// TIA Portal V20 export
// export: Created 2026-10-20T18:55:29.0460085Z, ExportSetting None, DisplayName Totally Integrated Automation Portal, DisplayVersion V20 Update 6, DisplayName TIA Portal Openness, DisplayVersion V20 Update 6, DisplayName TIA Portal Version Control Interface, DisplayVersion V20 Update 6, DisplayName SINAMICS Startdrive Advanced, DisplayVersion V20 SP1, DisplayName SINAMICS Startdrive G130, G150, S120, S150, SINAMICS MV, G220, S200, S210, DisplayVersion V20 SP1, DisplayName SINAMICS Startdrive G110M, G120, G120C, G120D, G120P, G115D, DisplayVersion V20 SP1, DisplayName STEP 7 Professional, DisplayVersion V20 Update 6, DisplayName STEP 7 Safety, DisplayVersion V20 Update 2, DisplayName WinCC Basic/Comfort/Advanced, DisplayVersion V20 Update 6, DisplayName WinCC Unified, DisplayVersion V20 Update 6
VAR_GLOBAL   // PLC tag table "IO_VFDs_5"
   C5103_StatusWord AT %IW2762 : Word;
   C5103_ActualCurrent AT %IW2766 : Word;
   C5102_ActualSpeed AT %IW2752 : Word;
   C5102_ActualCurrent AT %IW2754 : Word;
   C5104_StatusWord AT %IW2774 : Word;
   C5101_ControlWord AT %QW1349 : Word;
   VTD5_ActualCurrent AT %IW1630 : Word;
   C5107_ActualSpeed AT %IW2812 : Word;
   C5108_StatusWord AT %IW2822 : Word;
   CVTD5_ActualSpeed AT %IW2728 : Word;
   C5106_ControlWord AT %QW1472 : Word;
   C5105_ControlWord AT %QW1468 : Word;
   C5103_ActualSpeed AT %IW2764 : Word;
   C5108_MainSetpoint AT %QW1488 : Word;
   C5108_ControlWord AT %QW1486 : Word;
   C5103_ControlWord AT %QW1460 : Word;
   C5106_StatusWord AT %IW2798 : Word;
   C5106_ActualSpeed AT %IW2800 : Word;
   CVTD5_ActualCurrent AT %IW2730 : Word;
   C5104_ActualCurrent AT %IW2778 : Word;
   C5102_StatusWord AT %IW2750 : Word;
   C5105_ActualCurrent AT %IW2790 : Word;
   C5104_ControlWord AT %QW1464 : Word;
   C5101_StatusWord AT %IW2738 : Word;
   C5101_MainSetpoint AT %QW1351 : Word;
   C5107_ActualCurrent AT %IW2814 : Word;
   C5106_ActualCurrent AT %IW2802 : Word;
   C5101_ActualCurrent AT %IW2742 : Word;
   C5108_ActualSpeed AT %IW2824 : Word;
   C5103_MainSetpoint AT %QW1462 : Word;
   C5104_MainSetpoint AT %QW1466 : Word;
   C5106_MainSetpoint AT %QW1474 : Word;
   C5107_StatusWord AT %IW2810 : Word;
   C5105_MainSetpoint AT %QW1470 : Word;
   C5107_MainSetpoint AT %QW1484 : Word;
   CVTD5_MainSetpoint AT %QW1347 : Word;
   C5102_MainSetpoint AT %QW1355 : Word;
   C5108_ActualCurrent AT %IW2826 : Word;
   VTD5_StatusWord AT %IW1626 : Word;
   C5105_StatusWord AT %IW2786 : Word;
   CVTD5_StatusWord AT %IW2726 : Word;
   C5102_ControlWord AT %QW1353 : Word;
   C5101_ActualSpeed AT %IW2740 : Word;
   CVTD5_ControlWord AT %QW1345 : Word;
   C5105_ActualSpeed AT %IW2788 : Word;
   C5107_ControlWord AT %QW1482 : Word;
   C5104_ActualSpeed AT %IW2776 : Word;
   VTD5_ActualSpeed AT %IW1628 : Word;
   C5101_ActualTorque AT %IW2744 : Word;
   C5106_ActualTorque AT %IW2804 : Word;
   C5108_ActualTorque AT %IW2828 : Word;
   C5104_ActualTorque AT %IW2780 : Word;
   VTD5_ActualTorque AT %IW1632 : Word;
   C5107_ActualTorque AT %IW2816 : Word;
   C5103_ActualTorque AT %IW2768 : Word;
   C5102_ActualTorque AT %IW2756 : Word;
   CVTD5_ActualTorque AT %IW2732 : Word;
   C5105_ActualTorque AT %IW2792 : Word;
   VTD5_ControlWord AT %QW1341 : Word;
   VTD5_AccFactor AT %QW1509 : Word;
   VTD5_MainSetpoint AT %QW1343 : Word;
END_VAR
